DATA_BLOCK "FRK_Diagnostics"
{ S7_Optimized_Access := 'TRUE' }
VERSION : 0.1
NON_RETAIN
VAR
    Samples {ExternalAccessible := 'False'; ExternalVisible := 'False'; ExternalWritable := 'False'} : Array[1..7] of "FRK_DiagSample";
    Empty {ExternalAccessible := 'False'; ExternalVisible := 'False'; ExternalWritable := 'False'} : "FRK_DiagSummary";
END_VAR
BEGIN
END_DATA_BLOCK
